Fanuc KAREL source: kt00098.KL

-- PROVISIONAL review KL for V1013-1; original PC SHA256 ecd11d3c81630e7c26e100d2c434986d623f95f9d883223f45ee8f84e648d572
-- Incomplete behavior may be omitted. Consult companion uncertainty JSON. Do not deploy.
PROGRAM KT00098
%NOLOCKGROUP
VAR
  I1 : INTEGER
  I2 : INTEGER
  OUT : REAL
BEGIN
  -- UNRESOLVED_PC offsets 5-16; opcodes 2E,23
  -- UNRESOLVED_PC offsets 21-32; opcodes 2E,23
  -- UNRESOLVED_PC offsets 37-48; opcodes 2E,23
  -- UNRESOLVED_PC offsets 53-64; opcodes 2E,23
  -- UNRESOLVED_PC offsets 69-92; opcodes 21,21,64,29,64,29,6C,23
  -- UNRESOLVED_PC offsets 97-101; opcodes 7F
END KT00098
